(* IEC 61131-3 sources: gemelo-digital-planta/planta-clasificacion-gemelo-digital/plc-codesys, 2 files *)

(* ---- variables_globales.st ---- *)
(* =============================================================================
   variables_globales.st
   Proyecto : Planta Virtual de Clasificación Gobernada por PLC
   Norma    : IEC 61131-3:2013 · Texto Estructurado
   Contrato : config_modbus_slave.json v1.2.0 (4 tablas Modbus TCP: Coils 0..9,
              Discrete Inputs 0..10, Holding Registers 0..3, Input Registers 0..7;
              retrocompatible con las direcciones 0..6 de v1.1.0)
   Contiene : 4 objetos CODESYS a crear por separado en el árbol POU:
              [1] DUT  E_EstadoClasificador   (Enumeración de estados S0..S7)
              [2] DUT  E_ModoRuteo            (Enumeración de modos de ruteo)
              [3] GVL  GVL_IO                 (Imagen de proceso %IX, %QX, %MW, %IW)
              [4] GVL  GVL_Param              (Constantes de proceso por defecto)
   ============================================================================= *)

(* ------------------------------------------------------------------ [1] DUT -- *)
(* Estados S0..S7 de la máquina de Moore (docs/01 §3.1; S6 y S7 en v1.2.0).      *)
{attribute 'qualified_only'}
{attribute 'strict'}
{attribute 'to_string'}
TYPE E_EstadoClasificador :
(
    REPOSO                  := 0,   (* S0 · estado seguro de referencia, F = {S0} *)
    EN_MARCHA_ESPERA        := 1,   (* S1 · cinta activa esperando paquete en %IX0.3 *)
    CLASIFICANDO_RUTA_A     := 2,   (* S2 · evacuando hacia salida A hasta %IX0.7 *)
    CLASIFICANDO_RUTA_B     := 3,   (* S3 · evacuando hacia salida B hasta %IX1.0 *)
    PARADA_EMERGENCIA       := 4,   (* S4 · seta enclavada; requiere rearme consciente *)
    ESPERANDO_CAMBIO_ESTIBA := 5,   (* S5 · estiba A o B no disponible (llena o en cambio) *)
    FALLA_ATASCO            := 6,   (* S6 · watchdog TON vencido sin confirmar %IX0.7/%IX1.0 *)
    INSPECCION_NO_READ      := 7    (* S7 · código ilegible (SKU 99); espera asignación manual *)
) INT;
END_TYPE

(* ------------------------------------------------------------------ [2] DUT -- *)
{attribute 'qualified_only'}
{attribute 'strict'}
TYPE E_ModoRuteo :
(
    MANUAL        := 0,   (* Decide con %IX0.4 Selector_Destino *)
    AUTO_ESCANER  := 1,   (* Decide con %MW1 HR_SKU_Escaneado (1=A, 2=B, 99=NO_READ) *)
    AUTO_BALANCEO := 2    (* Alterna/balancea automáticamente en el PLC entre A y B *)
) UINT;
END_TYPE

(* ------------------------------------------------------------------ [3] GVL -- *)
(* Imagen de proceso. Las direcciones AT coinciden 1:1 con el esclavo Modbus:    *)
(*   Coils 0..9             -> %IX0.0..%IX1.1  (escritas por el maestro, FC05/15)*)
(*   Discrete Inputs 0..10  -> %QX0.0..%QX1.2  (leídas por el maestro, FC02)     *)
(*   Holding Registers 0..3 -> %MW0..%MW3      (leídos/escritos, FC03/FC06)      *)
(*   Input Registers 0..7   -> %IW0..%IW7      (telemetría PLC, FC04)            *)
{attribute 'qualified_only'}
VAR_GLOBAL
    (* Entradas discretas al PLC (%IX · Coils 0..9) ---------------------------- *)
    Marcha               AT %IX0.0 : BOOL;  (* Coil 0 · pulsador NA momentáneo         *)
    Parada               AT %IX0.1 : BOOL;  (* Coil 1 · pulsador momentáneo, prioridad *)
    Emergencia           AT %IX0.2 : BOOL;  (* Coil 2 · TRUE = emergencia activa       *)
    Sensor_Entrada       AT %IX0.3 : BOOL;  (* Coil 3 · fotocelda pórtico escáner      *)
    Selector_Destino     AT %IX0.4 : BOOL;  (* Coil 4 · FALSE = Ruta A, TRUE = Ruta B  *)
    Estiba_Llena_A       AT %IX0.5 : BOOL;  (* Coil 5 · estiba A no disponible         *)
    Estiba_Llena_B       AT %IX0.6 : BOOL;  (* Coil 6 · estiba B no disponible         *)
    Sensor_Salida_A      AT %IX0.7 : BOOL;  (* Coil 7 · fotocelda descarga salida A    *)
    Sensor_Salida_B      AT %IX1.0 : BOOL;  (* Coil 8 · fotocelda descarga salida B    *)
    Atasco_Planta        AT %IX1.1 : BOOL;  (* Coil 9 · atasco físico en banda activa  *)

    (* Salidas discretas del PLC (%QX · Discrete Inputs 0..10) ----------------- *)
    Motor_Cinta_Entrada  AT %QX0.0 : BOOL;  (* DI 0  · contactor banda principal       *)
    Actuador_Desviador   AT %QX0.1 : BOOL;  (* DI 1  · electroválvula 5/2 (TRUE = B)   *)
    Motor_Cinta_Salida_A AT %QX0.2 : BOOL;  (* DI 2  · contactor banda salida A        *)
    Motor_Cinta_Salida_B AT %QX0.3 : BOOL;  (* DI 3  · contactor banda salida B        *)
    Baliza_Alarma        AT %QX0.4 : BOOL;  (* DI 4  · torreta roja (S4 o S6)          *)
    Heartbeat_Out        AT %QX0.5 : BOOL;  (* DI 5  · onda cuadrada supervisión ~1 Hz *)
    Senal_Cambio_Estiba  AT %QX0.6 : BOOL;  (* DI 6  · torreta ámbar (S5 o S7)         *)
    Stopper_Admision     AT %QX0.7 : BOOL;  (* DI 7  · tope neumático indexador cola   *)
    Alarma_Atasco        AT %QX1.0 : BOOL;  (* DI 8  · falla de watchdog de atasco S6  *)
    Aviso_NoRead         AT %QX1.1 : BOOL;  (* DI 9  · pausa inspección NO_READ S7     *)
    Baliza_Verde         AT %QX1.2 : BOOL;  (* DI 10 · torreta verde operación normal  *)

    (* Registros de mantenimiento (%MW · Holding Registers 0..3, FC03/FC06) ---- *)
    HR_Modo_Ruteo          AT %MW0 : UINT := 0;    (* 0=Manual, 1=Escáner, 2=Balanceo *)
    HR_SKU_Escaneado       AT %MW1 : UINT := 0;    (* 0=Sin dato, 1=SKU_A, 2=SKU_B, 99=NO_READ *)
    HR_Modo_Watchdog       AT %MW2 : UINT := 0;    (* 0=Clásico/Señal, 1=Lazo cerrado estricto *)
    HR_Tiempo_Watchdog_Ms  AT %MW3 : UINT := 4000; (* PT del watchdog en ms (1000..15000) *)

    (* Registros de entrada (%IW · Input Registers 0..7, FC04) ----------------- *)
    IR_Estado_FSM          AT %IW0 : UINT;  (* Código numérico E_EstadoClasificador 0..7 *)
    IR_Codigo_Falla        AT %IW1 : UINT;  (* 0=OK, 1=EMERG, 2=ESTIBA, 3=ATASCO, 4=NOREAD, 5=COHERENCIA *)
    IR_Paquetes_A          AT %IW2 : UINT;  (* Contador acumulado Ruta A                *)
    IR_Paquetes_B          AT %IW3 : UINT;  (* Contador acumulado Ruta B                *)
    IR_Atascos             AT %IW4 : UINT;  (* Contador acumulado de atascos            *)
    IR_NoRead              AT %IW5 : UINT;  (* Contador acumulado de lecturas NO_READ   *)
    IR_Tiempo_Clasif_Ms    AT %IW6 : UINT;  (* Tiempo transcurrido ET del TON (ms)      *)
    IR_Ultimo_SKU          AT %IW7 : UINT;  (* Último SKU evaluado en el túnel lector   *)
END_VAR

(* ------------------------------------------------------------------ [4] GVL -- *)
{attribute 'qualified_only'}
VAR_GLOBAL CONSTANT
    T_HEARTBEAT     : TIME := T#500MS;  (* PT de Heartbeat_Timer (semiperiodo)          *)
    T_CLASIFICACION : TIME := T#4S;     (* T_clas / Watchdog por defecto (docs/01 §3.2) *)
END_VAR

(* ---- logica_clasificador_fsm.st ---- *)
(* =============================================================================
   logica_clasificador_fsm.st
   Proyecto : Planta Virtual de Clasificación Gobernada por PLC
   Norma    : IEC 61131-3:2013 · Texto Estructurado
   Modelo   : Máquina de Moore M = (S, Σ, Λ, δ, λ, s0, F) — Contrato v1.2.0
   Contiene : 3 POU a crear por separado (Agregar objeto > POU):
              [1] FB_Heartbeat        (Bloque de función)
              [2] FB_ClasificadorFSM  (Bloque de función)
              [3] PLC_PRG             (Programa · asignado a MainTask, cíclica T#10MS)
   Depende  : variables_globales.st (E_EstadoClasificador, E_ModoRuteo, GVL_IO, GVL_Param)
   ============================================================================= *)

(* ========================================================= [1] FB_Heartbeat == *)
FUNCTION_BLOCK FB_Heartbeat
VAR_INPUT
    tSemiperiodo : TIME := T#500MS;
END_VAR
VAR_OUTPUT
    xPulso : BOOL;                 (* h *)
END_VAR
VAR
    Heartbeat_Timer : TON;         (* nombre exigido por la especificación *)
END_VAR

Heartbeat_Timer(IN := NOT Heartbeat_Timer.Q, PT := tSemiperiodo);
IF Heartbeat_Timer.Q THEN
    xPulso := NOT xPulso;
END_IF
END_FUNCTION_BLOCK

(* =================================================== [2] FB_ClasificadorFSM == *)
(* Orden de evaluación por ciclo de scan k:                                     *)
(*   (a) detección de flancos m↑, s↑, sA↑, sB↑ (R_TRIG, siempre — propiedad P4) *)
(*   (b) t = TON_Clasif(IN := s(k) ∈ {S2,S3}, PT := tClasificacion).Q            *)
(*   (c) s(k+1) = δ(s(k), σ(k))                                                 *)
(*       Prioridad: Emergencia ≻ Estiba no disponible ≻ Parada ≻ Proceso         *)
(*   (d) Q(k) = λ(s(k+1))              salida de Moore inyectiva                *)
(*   (e) diagnóstico de invariantes P2/P3 y código de falla                     *)
FUNCTION_BLOCK FB_ClasificadorFSM
VAR_INPUT
    xMarcha         : BOOL;    (* m  · %IX0.0 *)
    xParada         : BOOL;    (* p  · %IX0.1 *)
    xEmergencia     : BOOL;    (* e  · %IX0.2 TRUE = activa *)
    xSensor         : BOOL;    (* s  · %IX0.3 fotocelda entrada *)
    xSelectorB      : BOOL;    (* d  · %IX0.4 FALSE = A, TRUE = B *)
    xEstibaLlenaA   : BOOL;    (* ℓA · %IX0.5 *)
    xEstibaLlenaB   : BOOL;    (* ℓB · %IX0.6 *)
    xSensorSalidaA  : BOOL;    (* sA · %IX0.7 fotocelda salida A *)
    xSensorSalidaB  : BOOL;    (* sB · %IX1.0 fotocelda salida B *)
    xAtascoPlanta   : BOOL;    (* j  · %IX1.1 condición física de atasco *)
    uiModoRuteo     : UINT := 0;    (* %MW0: 0=Manual, 1=Escáner, 2=Balanceo *)
    uiSkuEscaneado  : UINT := 0;    (* %MW1: 0=Sin dato, 1=A, 2=B, 99=NO_READ *)
    uiModoWatchdog  : UINT := 0;    (* %MW2: 0=Clásico/Atasco, 1=Estricto lazo cerrado *)
    tClasificacion  : TIME := T#4S; (* %MW3 / GVL_Param.T_CLASIFICACION *)
END_VAR
VAR_OUTPUT
    xCintaEntrada      : BOOL; (* Q0  · %QX0.0 *)
    xDesviador         : BOOL; (* Q1  · %QX0.1 *)
    xCintaSalidaA      : BOOL; (* Q2  · %QX0.2 *)
    xCintaSalidaB      : BOOL; (* Q3  · %QX0.3 *)
    xBaliza            : BOOL; (* Q4  · %QX0.4 *)
    xSenalCambioEstiba : BOOL; (* Q6  · %QX0.6 *)
    xStopperAdmision   : BOOL; (* Q7  · %QX0.7 tope indexador de admisión *)
    xAlarmaAtasco      : BOOL; (* Q8  · %QX1.0 falla de watchdog *)
    xAvisoNoRead       : BOOL; (* Q9  · %QX1.1 pausa inspección NO_READ *)
    xBalizaVerde       : BOOL; (* Q10 · %QX1.2 operación normal *)
    eEstado            : E_EstadoClasificador := E_EstadoClasificador.REPOSO;
    xFallaCoherencia   : BOOL;
    uiCodigoFalla      : UINT := 0;
    udiPaquetesA       : UDINT := 0;
    udiPaquetesB       : UDINT := 0;
    udiAtascos         : UDINT := 0;
    udiNoRead          : UDINT := 0;
    uiTiempoClasifMs   : UINT := 0;
    uiUltimoSku        : UINT := 0;
END_VAR
VAR
    rtMarcha           : R_TRIG;
    rtSensor           : R_TRIG;
    rtSalidaA          : R_TRIG;
    rtSalidaB          : R_TRIG;
    TON_Clasif         : TON;
    xTurnoBalanceoB    : BOOL := FALSE;
    xIrRutaB           : BOOL := FALSE;
END_VAR

(* (a) Flancos ascendentes: evaluados en todo ciclo (P4) *)
rtMarcha(CLK := xMarcha);
rtSensor(CLK := xSensor);
rtSalidaA(CLK := xSensorSalidaA);
rtSalidaB(CLK := xSensorSalidaB);

(* (b) Temporizador / Watchdog de clasificación sobre el estado vigente *)
TON_Clasif(IN := (eEstado = E_EstadoClasificador.CLASIFICANDO_RUTA_A)
              OR (eEstado = E_EstadoClasificador.CLASIFICANDO_RUTA_B),
           PT := tClasificacion);
uiTiempoClasifMs := TIME_TO_UINT(TON_Clasif.ET);

(* (c) Función de transición δ *)
IF xEmergencia THEN                                             (* T1 · ∀s → S4 *)
    eEstado := E_EstadoClasificador.PARADA_EMERGENCIA;
ELSIF (xEstibaLlenaA OR xEstibaLlenaB)
      AND eEstado <> E_EstadoClasificador.PARADA_EMERGENCIA
      AND eEstado <> E_EstadoClasificador.FALLA_ATASCO THEN     (* T9 · S0..S3, S7 → S5 *)
    eEstado := E_EstadoClasificador.ESPERANDO_CAMBIO_ESTIBA;
ELSE
    CASE eEstado OF
    E_EstadoClasificador.REPOSO:
        IF NOT xParada AND rtMarcha.Q THEN                      (* T2 *)
            eEstado := E_EstadoClasificador.EN_MARCHA_ESPERA;
        END_IF

    E_EstadoClasificador.EN_MARCHA_ESPERA:
        IF xParada THEN                                         (* T3 *)
            eEstado := E_EstadoClasificador.REPOSO;
        ELSIF rtSensor.Q THEN                                   (* Muestreo de destino en s↑ (P5) *)
            IF uiModoRuteo = 1 THEN                             (* Modo 1: AUTO_ESCANER *)
                uiUltimoSku := uiSkuEscaneado;
                IF uiSkuEscaneado = 99 THEN                     (* T13 · Código ilegible → S7 *)
                    eEstado := E_EstadoClasificador.INSPECCION_NO_READ;
                    udiNoRead := udiNoRead + 1;
                ELSIF uiSkuEscaneado = 2 THEN
                    eEstado := E_EstadoClasificador.CLASIFICANDO_RUTA_B;
                    udiPaquetesB := udiPaquetesB + 1;
                ELSE
                    eEstado := E_EstadoClasificador.CLASIFICANDO_RUTA_A;
                    udiPaquetesA := udiPaquetesA + 1;
                END_IF
            ELSIF uiModoRuteo = 2 THEN                          (* Modo 2: AUTO_BALANCEO *)
                xIrRutaB := xTurnoBalanceoB;
                xTurnoBalanceoB := NOT xTurnoBalanceoB;
                uiUltimoSku := SEL(xIrRutaB, 1, 2);
                IF xIrRutaB THEN
                    eEstado := E_EstadoClasificador.CLASIFICANDO_RUTA_B;
                    udiPaquetesB := udiPaquetesB + 1;
                ELSE
                    eEstado := E_EstadoClasificador.CLASIFICANDO_RUTA_A;
                    udiPaquetesA := udiPaquetesA + 1;
                END_IF
            ELSE                                                (* Modo 0: MANUAL (%IX0.4) *)
                uiUltimoSku := SEL(xSelectorB, 1, 2);
                IF xSelectorB THEN                              (* T5 *)
                    eEstado := E_EstadoClasificador.CLASIFICANDO_RUTA_B;
                    udiPaquetesB := udiPaquetesB + 1;
                ELSE                                            (* T4 *)
                    eEstado := E_EstadoClasificador.CLASIFICANDO_RUTA_A;
                    udiPaquetesA := udiPaquetesA + 1;
                END_IF
            END_IF
        END_IF

    E_EstadoClasificador.CLASIFICANDO_RUTA_A:
        IF xParada THEN                                         (* T7 *)
            eEstado := E_EstadoClasificador.REPOSO;
        ELSIF rtSalidaA.Q AND NOT xAtascoPlanta THEN            (* T6a · Cierre de lazo en salida A *)
            eEstado := E_EstadoClasificador.EN_MARCHA_ESPERA;
        ELSIF TON_Clasif.Q THEN
            IF xAtascoPlanta OR (uiModoWatchdog = 1) THEN       (* T11 · Watchdog vencido sin descarga → S6 *)
                eEstado := E_EstadoClasificador.FALLA_ATASCO;
                udiAtascos := udiAtascos + 1;
            ELSE                                                (* T6 · Lazo abierto clásico *)
                eEstado := E_EstadoClasificador.EN_MARCHA_ESPERA;
            END_IF
        END_IF

    E_EstadoClasificador.CLASIFICANDO_RUTA_B:
        IF xParada THEN                                         (* T7 *)
            eEstado := E_EstadoClasificador.REPOSO;
        ELSIF rtSalidaB.Q AND NOT xAtascoPlanta THEN            (* T6b · Cierre de lazo en salida B *)
            eEstado := E_EstadoClasificador.EN_MARCHA_ESPERA;
        ELSIF TON_Clasif.Q THEN
            IF xAtascoPlanta OR (uiModoWatchdog = 1) THEN       (* T11 · Watchdog vencido sin descarga → S6 *)
                eEstado := E_EstadoClasificador.FALLA_ATASCO;
                udiAtascos := udiAtascos + 1;
            ELSE                                                (* T6 · Lazo abierto clásico *)
                eEstado := E_EstadoClasificador.EN_MARCHA_ESPERA;
            END_IF
        END_IF

    E_EstadoClasificador.PARADA_EMERGENCIA:
        IF xParada THEN                                         (* T8 · Rearme consciente *)
            eEstado := E_EstadoClasificador.REPOSO;
        END_IF

    E_EstadoClasificador.ESPERANDO_CAMBIO_ESTIBA:
        eEstado := E_EstadoClasificador.REPOSO;                 (* T10 · exige Marcha (P7) *)

    E_EstadoClasificador.FALLA_ATASCO:
        IF xParada AND NOT xAtascoPlanta THEN                   (* T12 · Rearme tras despejar atasco *)
            eEstado := E_EstadoClasificador.REPOSO;
        END_IF

    E_EstadoClasificador.INSPECCION_NO_READ:
        IF xParada THEN                                         (* Cancelar a Reposo *)
            eEstado := E_EstadoClasificador.REPOSO;
        ELSIF rtMarcha.Q THEN                                   (* T14 · Operador asigna ruta A/B y confirma con Marcha *)
            IF xSelectorB THEN
                uiUltimoSku := 2;
                eEstado := E_EstadoClasificador.CLASIFICANDO_RUTA_B;
                udiPaquetesB := udiPaquetesB + 1;
            ELSE
                uiUltimoSku := 1;
                eEstado := E_EstadoClasificador.CLASIFICANDO_RUTA_A;
                udiPaquetesA := udiPaquetesA + 1;
            END_IF
        END_IF

    ELSE
        eEstado := E_EstadoClasificador.PARADA_EMERGENCIA;
    END_CASE
END_IF

(* (d) Función de salida λ (Moore): códigos inyectivos *)
xCintaEntrada      := (eEstado = E_EstadoClasificador.EN_MARCHA_ESPERA)
                   OR (eEstado = E_EstadoClasificador.CLASIFICANDO_RUTA_A)
                   OR (eEstado = E_EstadoClasificador.CLASIFICANDO_RUTA_B);
xDesviador         :=  eEstado = E_EstadoClasificador.CLASIFICANDO_RUTA_B;
xCintaSalidaA      :=  eEstado = E_EstadoClasificador.CLASIFICANDO_RUTA_A;
xCintaSalidaB      :=  eEstado = E_EstadoClasificador.CLASIFICANDO_RUTA_B;
xBaliza            := (eEstado = E_EstadoClasificador.PARADA_EMERGENCIA)
                   OR (eEstado = E_EstadoClasificador.FALLA_ATASCO);
xSenalCambioEstiba := (eEstado = E_EstadoClasificador.ESPERANDO_CAMBIO_ESTIBA)
                   OR (eEstado = E_EstadoClasificador.INSPECCION_NO_READ);
xStopperAdmision   := (eEstado = E_EstadoClasificador.CLASIFICANDO_RUTA_A)
                   OR (eEstado = E_EstadoClasificador.CLASIFICANDO_RUTA_B)
                   OR (eEstado = E_EstadoClasificador.INSPECCION_NO_READ)
                   OR (eEstado = E_EstadoClasificador.FALLA_ATASCO);
xAlarmaAtasco      :=  eEstado = E_EstadoClasificador.FALLA_ATASCO;
xAvisoNoRead       :=  eEstado = E_EstadoClasificador.INSPECCION_NO_READ;
xBalizaVerde       :=  xCintaEntrada;

(* (e) Invariantes P2/P3 y código de falla *)
xFallaCoherencia := (xCintaSalidaA AND xCintaSalidaB) OR (xDesviador XOR xCintaSalidaB);

IF xFallaCoherencia THEN
    uiCodigoFalla := 5;
ELSIF eEstado = E_EstadoClasificador.PARADA_EMERGENCIA THEN
    uiCodigoFalla := 1;
ELSIF eEstado = E_EstadoClasificador.ESPERANDO_CAMBIO_ESTIBA THEN
    uiCodigoFalla := 2;
ELSIF eEstado = E_EstadoClasificador.FALLA_ATASCO THEN
    uiCodigoFalla := 3;
ELSIF eEstado = E_EstadoClasificador.INSPECCION_NO_READ THEN
    uiCodigoFalla := 4;
ELSE
    uiCodigoFalla := 0;
END_IF
END_FUNCTION_BLOCK

(* ================================================================ [3] PLC_PRG == *)
PROGRAM PLC_PRG
VAR
    fbClasificador : FB_ClasificadorFSM;
    fbHeartbeat    : FB_Heartbeat;
    tWatchdog      : TIME;
END_VAR

fbHeartbeat(tSemiperiodo := GVL_Param.T_HEARTBEAT);

IF GVL_IO.HR_Tiempo_Watchdog_Ms >= 1000 AND GVL_IO.HR_Tiempo_Watchdog_Ms <= 15000 THEN
    tWatchdog := UINT_TO_TIME(GVL_IO.HR_Tiempo_Watchdog_Ms);
ELSE
    tWatchdog := GVL_Param.T_CLASIFICACION;
END_IF

fbClasificador(
    xMarcha        := GVL_IO.Marcha,
    xParada        := GVL_IO.Parada,
    xEmergencia    := GVL_IO.Emergencia,
    xSensor        := GVL_IO.Sensor_Entrada,
    xSelectorB     := GVL_IO.Selector_Destino,
    xEstibaLlenaA  := GVL_IO.Estiba_Llena_A,
    xEstibaLlenaB  := GVL_IO.Estiba_Llena_B,
    xSensorSalidaA := GVL_IO.Sensor_Salida_A,
    xSensorSalidaB := GVL_IO.Sensor_Salida_B,
    xAtascoPlanta  := GVL_IO.Atasco_Planta,
    uiModoRuteo    := GVL_IO.HR_Modo_Ruteo,
    uiSkuEscaneado := GVL_IO.HR_SKU_Escaneado,
    uiModoWatchdog := GVL_IO.HR_Modo_Watchdog,
    tClasificacion := tWatchdog);

(* Escritura de la imagen de salidas discretas %QX *)
GVL_IO.Motor_Cinta_Entrada  := fbClasificador.xCintaEntrada;
GVL_IO.Actuador_Desviador   := fbClasificador.xDesviador;
GVL_IO.Motor_Cinta_Salida_A := fbClasificador.xCintaSalidaA;
GVL_IO.Motor_Cinta_Salida_B := fbClasificador.xCintaSalidaB;
GVL_IO.Baliza_Alarma        := fbClasificador.xBaliza OR fbClasificador.xFallaCoherencia;
GVL_IO.Heartbeat_Out        := fbHeartbeat.xPulso;
GVL_IO.Senal_Cambio_Estiba  := fbClasificador.xSenalCambioEstiba;
GVL_IO.Stopper_Admision     := fbClasificador.xStopperAdmision;
GVL_IO.Alarma_Atasco        := fbClasificador.xAlarmaAtasco;
GVL_IO.Aviso_NoRead         := fbClasificador.xAvisoNoRead;
GVL_IO.Baliza_Verde         := fbClasificador.xBalizaVerde;

(* Escritura de los registros de entrada %IW (telemetría FC04) *)
GVL_IO.IR_Estado_FSM        := INT_TO_UINT(fbClasificador.eEstado);
GVL_IO.IR_Codigo_Falla      := fbClasificador.uiCodigoFalla;
GVL_IO.IR_Paquetes_A        := UDINT_TO_UINT(fbClasificador.udiPaquetesA);
GVL_IO.IR_Paquetes_B        := UDINT_TO_UINT(fbClasificador.udiPaquetesB);
GVL_IO.IR_Atascos           := UDINT_TO_UINT(fbClasificador.udiAtascos);
GVL_IO.IR_NoRead            := UDINT_TO_UINT(fbClasificador.udiNoRead);
GVL_IO.IR_Tiempo_Clasif_Ms  := fbClasificador.uiTiempoClasifMs;
GVL_IO.IR_Ultimo_SKU        := fbClasificador.uiUltimoSku;
END_PROGRAM
